(* IEC 61131-3 sources: 2026_Projet_YGO_ExcavatriceDragage/CODE_BACKUP/CODE_20260807_v0.5.25/JOYSTICK, 4 files *)

(* ---- ST_Joystick_AxisCmd.st ---- *)
(* ═══════════════════════════════════════════════════════════════
   🕹️ ST_Joystick_AxisCmd — Consigne d'axe normalisée (sortie FB_Joystick)
   ───────────────────────────────────────────────────────────────
   📄 Doc métier : DOC/AF_Partie-08_Fonction_Joystick_v2.0.md
                   DOC/AF_Partie-03_Contrats_Composants_v2.1.md
   🎯 4 champs exactement :
      - Enable    : Autorisation globale du pipeline
      - StartStop : RAMPE (TRUE = accélération, FALSE = décélération normale)
      - SpeedRef  : Consigne vitesse signée (-100.0 .. +100.0 %)
      - Direction : Sens d'axe (-1 = Rev, 0 = Neutre, +1 = Fwd)
   ═══════════════════════════════════════════════════════════════ *)

TYPE ST_Joystick_AxisCmd :
STRUCT
    Enable      : BOOL;   // Autorisation FB (FALSE = neutralisation, sorties coupées)
    StartStop   : BOOL;   // TRUE = rampe accélération, FALSE = rampe décélération normale
    SpeedRef    : REAL;   // Consigne vitesse SIGNÉE -100..+100 % (signe = sens, cohérent avec Direction)
    Direction   : INT;    // -1 = Rev, 0 = Neutre, +1 = Fwd
END_STRUCT
END_TYPE

(* ---- FB_AxisScale.st ---- *)
(* ═══════════════════════════════════════════════════════════════
   📐 FB_AxisScale — Mise à l'échelle d'un axe joystick Hall
   ───────────────────────────────────────────────────────────────
   📄 Extrait depuis le projet CODESYS (Device.export, JOYSTICK/)
   🎯 Normalise une valeur brute (0..10000) par rapport au neutre calibré
      et applique une zone morte en unités brutes (compte ADC, pas en %).
   Sortie : OutPct ∈ [-100.0 .. +100.0] (0.0 si dans la deadband)
   🔧 2026-08-07 (demande client) : Deadband (REAL, %) → DeadbandRaw (INT, compte brut 0..10000).
      Raison : plus simple à régler directement depuis le bruit mesuré au neutre (ex: ±200 sur le
      terrain → DeadbandRaw=300 avec marge), sans recalculer un % à chaque calibration.
   ═══════════════════════════════════════════════════════════════
   📄 Docs : DOC/AF_Partie-08_Fonction_Joystick_v2.0.md
*)

FUNCTION_BLOCK FB_AxisScale
VAR_INPUT
    /// Valeur brute (0..10000)
    RawIn   : INT;
    /// Point milieu calibré
    Neutral : INT;
    /// Zone morte en unités brutes (compte ADC, ex: 300 sur plage 0..10000)
    DeadbandRaw : INT;
END_VAR
VAR_OUTPUT
    /// Valeur finale (-100.0..100.0)
    OutPct : REAL;
END_VAR
VAR
    Delta : REAL;
END_VAR

IF RawIn >= Neutral THEN
    Delta := INT_TO_REAL(10000 - Neutral);
    IF Delta > 0.0 THEN
        OutPct := (INT_TO_REAL(RawIn - Neutral) / Delta) * 100.0;
    ELSE
        OutPct := 0.0;
    END_IF;
ELSE
    Delta := INT_TO_REAL(Neutral);
    IF Delta > 0.0 THEN
        OutPct := (INT_TO_REAL(RawIn - Neutral) / Delta) * 100.0;
    ELSE
        OutPct := 0.0;
    END_IF;
END_IF;

IF ABS(RawIn - Neutral) <= DeadbandRaw THEN
    OutPct := 0.0;
END_IF;

// 🛡️ Limitation de plage : une valeur brute hors plage nominale ne doit jamais
// produire une consigne supérieure à ±100 %. Ce garde-fou protège les
// consommateurs en aval, notamment la translation M3.
OutPct := LIMIT(-100.0, OutPct, 100.0);

(* ---- FB_Filter_PT1.st ---- *)
(* ═══════════════════════════════════════════════════════════════
   🔁 FB_Filter_PT1 — Filtre passe-bas premier ordre (PT1 numérique)
   ───────────────────────────────────────────────────────────────
   📄 Extrait depuis le projet CODESYS (Device.export, JOYSTICK/)
   🎯 Filtre exponentiel discret : y[k] = α·x[k] + (1-α)·y[k-1]
      où α = CycleTimeS / (T + CycleTimeS), T = TimeConst en secondes.
   ⚠️ Si TimeConst = 0 ou CycleTimeS = 0, sortie = entrée (pass-through).
   ═══════════════════════════════════════════════════════════════
   📄 Docs : DOC/AF_Partie-08_Fonction_Joystick_v2.0.md
*)

FUNCTION_BLOCK FB_Filter_PT1
VAR_INPUT
    /// Consigne brute entrée
    ValueIn    : REAL;
    /// Constante de temps du filtre
    TimeConst  : TIME;
    /// Temps de cycle réel en secondes
    CycleTimeS : REAL;
END_VAR
VAR_OUTPUT
    /// Consigne filtrée sortie
    ValueOut : REAL;
END_VAR
VAR
    T     : REAL;
    Alpha : REAL;
END_VAR

T := TIME_TO_REAL(TimeConst) / 1000.0; // ms → s

IF T <= 0.0 OR CycleTimeS <= 0.0 THEN
    ValueOut := ValueIn;
ELSE
    Alpha    := CycleTimeS / (T + CycleTimeS);
    ValueOut := Alpha * ValueIn + (1.0 - Alpha) * ValueOut;
END_IF;

(* ---- FB_Joystick.st ---- *)
(* ═══════════════════════════════════════════════════════════════
   🕹️ FB_Joystick — Acquisition & traitement Hall (Homme-mort ISO 13850)
   ───────────────────────────────────────────────────────────────
   📄 Doc métier : DOC/AF_Partie-08_Fonction_Joystick_v2.0.md
                   DOC/AF_Partie-03_Contrats_Composants_v2.1.md
   🎯 Rôle : Acquisition 2 axes Hall + bouton homme-mort normatif.
      Pipeline par axe : FB_AxisScale → FB_Filter_PT1 → Homme-Mort → ST_Joystick_AxisCmd.
      Les rampes d'accélération/décélération sont gérées exclusivement par les
      FB de mouvement aval (FB_Winch, FB_Translation), hors de ce bloc.
    🔒 Bouton homme-mort :
       - Armement au neutre strict (ScaleX/Y.OutPct = 0.0).
       - Consentement au démarrage : mouvement libre SANS surveillance du bouton
         (défaut, DeadmanReconfEnable := FALSE). Optionnel : reconfirmation périodique
         en mouvement (délai DeadmanRearmTimeout) si DeadmanReconfEnable := TRUE.
       - Désarmement sur maintien au neutre (durée NeutralHoldTime) + gate/mode/fin benne.
   📤 Produit AxisCmdX, AxisCmdY, et signaux de diagnostic/miroir.
   ═══════════════════════════════════════════════════════════════ *)

// === DECLARATION (à coller dans la partie déclaration du POU FB_Joystick) ===

FUNCTION_BLOCK FB_Joystick
VAR_INPUT
    Enable          : BOOL;       // Active la logique
    Reset           : BOOL;       // Acquittement défaut
    PowerContactorEngaged : BOOL;       // Conditions globales OK (chaîne AU réarmée)
    Mode            : E_Mode;     // Changement de mode désarme le homme-mort
    BenneBusy       : BOOL;       // Fin de cycle benne (front descendant) désarme le homme-mort
    PreserveArmingAfterBucket : BOOL; // TRUE uniquement pendant fermeture ExtractionSequence : enchaînement palier 1 autorisé
    BusCanOpenOP    : ST_Diag_Device;       // État présence nœud CAN
    JoystickOP      : ST_Diag_Device;       // Mode esclave CANopen actif
    RawX            : INT;        // Valeur brute axe X
    RawY            : INT;        // Valeur brute axe Y
    RawButton       : BOOL;       // État brut bouton
    BtnCalibrate    : BOOL;       // Demande de recalage neutre
    InvertX         : BOOL := FALSE;
    InvertY         : BOOL := FALSE;
    DeadbandRaw     : INT := 300;    // 🔧 2026-08-07 (demande client) : zone morte en compte brut ADC (0..10000), remplace l'ancien % — mesure terrain bruit neutre ±200, marge à ±300
    FilterTime      : TIME := TIME#0ms;
    DeadmanRearmTimeout : TIME := T#10S; // Délai max entre 2 appuis en mouvement (si reconfirmation activée)
    NeutralHoldTime     : TIME := T#100MS; // Temps continu au neutre avant désarmement (100 ms)
    DeadmanArmHoldTime  : TIME := T#100MS; // 🆕 2026-08-07 : Temps d'appui continu avant armement (indépendant position axes)
    DeadmanArmGraceTime : TIME := T#3S;    // 🆕 2026-08-07 : Délai après armement avant que le désarmement "neutre tenu" (NeutralHoldTime) puisse s'appliquer — laisse le temps de sortir de la zone morte après un appui au centre
    DeadmanReconfEnable : BOOL := FALSE; // 🆕 2026-08-03 : FALSE = bouton = consentement au démarrage (mouvement libre, défaut cible) ; TRUE = reconfirmation périodique en mouvement (comportement historique)
END_VAR
VAR_OUTPUT
    Ready           : BOOL;       // Prêt à commuter
    Busy            : BOOL;       // Traitement en cours
    Done            : BOOL;       // Données valides dispo
    Error           : BOOL;       // Présence anomalie
    ErrorId         : WORD;       // bit0: "Échec calibration Joystick" - Valeurs RawX/Y hors plage lors du recalage
    AxisCmdX        : ST_Joystick_AxisCmd; // Sortie normalisée X
    AxisCmdY        : ST_Joystick_AxisCmd; // Sortie normalisée Y
    Button          : BOOL;       // Bouton filtré
    NeutralXAct     : INT;        // Point neutre X actuel pour IHM/Test
    NeutralYAct     : INT;        // Point neutre Y actuel pour IHM/Test
    // 🆕 Miroirs directs (maintenance) — mêmes valeurs que AxisCmdX/Y.SpeedRef/.Direction,
    // exposés à plat pour lecture immédiate en vue instance CODESYS (pas de dépliage struct).
    SpeedXPct       : REAL;       // Consigne vitesse axe X en % SIGNÉE (-100..+100), miroir AxisCmdX.SpeedRef
    DirectionX      : INT;        // Sens axe X (-1=Rev/0=Neutre/+1=Fwd), miroir AxisCmdX.Direction
    SpeedYPct       : REAL;       // Consigne vitesse axe Y en % SIGNÉE (-100..+100), miroir AxisCmdY.SpeedRef
    DirectionY      : INT;        // Sens axe Y (-1=Rev/0=Neutre/+1=Fwd), miroir AxisCmdY.Direction
    DeadmanArmed    : BOOL;       // 🆕 Geste armé (bouton appuyé au neutre) — IHM/diagnostic
    AtNeutral       : BOOL;       // 🆕 2026-08-07 : TRUE si les 2 axes sont en zone morte (position centrale) — IHM/diagnostic
END_VAR
VAR_IN_OUT
    NeutralXMem     : INT; // Point neutre X persistant global
    NeutralYMem     : INT; // Point neutre Y persistant global
END_VAR
VAR
    CycleTimeCalc   : FB_CycleTime;
    ScaleX          : FB_AxisScale;
    ScaleY          : FB_AxisScale;
    FilterX         : FB_Filter_PT1;
    FilterY         : FB_Filter_PT1;
    CmdXVal         : REAL;
    CmdYVal         : REAL;
    LastCalibrate   : BOOL;
    ResetEdge       : R_TRIG;
    DeadmanEdge     : R_TRIG;
    DeadmanTimer    : TON;
    NeutralHoldTimer: TON;
    DeadmanArmTimer : TON;
    DeadmanArmPending : BOOL;
    DeadmanArmGraceTimer : TON;
    LastMode        : E_Mode;
    BenneBusyFallEdge : F_TRIG;
END_VAR

// === IMPLEMENTATION (à coller dans le corps ST du POU FB_Joystick) ===

// 🛑 1. GATE (Sécurités et coupures prioritaires)
IF NOT Enable OR NOT PowerContactorEngaged OR NOT BusCanOpenOP.Operational OR NOT JoystickOP.Operational THEN
    Ready := FALSE; Busy := FALSE; Done := FALSE;
    AxisCmdX.Enable := FALSE; AxisCmdX.StartStop := FALSE; AxisCmdX.SpeedRef := 0.0; AxisCmdX.Direction := 0;
    AxisCmdY.Enable := FALSE; AxisCmdY.StartStop := FALSE; AxisCmdY.SpeedRef := 0.0; AxisCmdY.Direction := 0;
    SpeedXPct := 0.0; DirectionX := 0;
    SpeedYPct := 0.0; DirectionY := 0;
    Button := FALSE;
    AtNeutral := TRUE;   // 🆕 2026-08-07 — pas de commande possible pendant la neutralisation
    DeadmanArmed := FALSE;   // 🆕 Désarmé sur toute neutralisation — nouvel appui au neutre exigé
    DeadmanArmPending := FALSE;   // 🆕 2026-08-07 — annule toute tentative d'armement en cours
    DeadmanTimer(IN := FALSE, PT := DeadmanRearmTimeout);   // 🆕 2026-07-03decies — pas d'accumulation à froid
    NeutralHoldTimer(IN := FALSE, PT := NeutralHoldTime);   // 🆕 2026-07-03duodecies — idem
    DeadmanArmTimer(IN := FALSE, PT := DeadmanArmHoldTime);   // 🆕 2026-08-07 — idem
    DeadmanArmGraceTimer(IN := FALSE, PT := DeadmanArmGraceTime);   // 🆕 2026-08-07 — idem
    NeutralXAct := NeutralXMem;
    NeutralYAct := NeutralYMem;
    LastMode := Mode;   // 🆕 REX 2026-07-08 — pas de faux changement détecté à la réactivation
    RETURN;
END_IF;

Ready := TRUE; Busy := TRUE;

// 🔑 2. RESET DÉFAUT (front + cause disparue, Partie3 §5)
ResetEdge(CLK := Reset);
IF ResetEdge.Q AND (RawX >= 2000 AND RawX <= 8000 AND RawY >= 2000 AND RawY <= 8000) THEN
    ErrorId := ErrorId AND 16#FFFE;
END_IF;

// 📥 3. ACQUISITION TIMING & BOUTON
CycleTimeCalc();
Button := RawButton;

// 🎯 4. CALIBRATION DYNAMIQUE (Zone RETAIN)
IF BtnCalibrate AND NOT LastCalibrate THEN
    IF RawX >= 2000 AND RawX <= 8000 AND RawY >= 2000 AND RawY <= 8000 THEN
        NeutralXMem := RawX;
        NeutralYMem := RawY;
    ELSE
        // Un seul bit pour une seule cause (Partie3 §3)
        ErrorId := ErrorId OR 16#0001;
    END_IF;
END_IF;
Error := (ErrorId <> 16#0000);
LastCalibrate := BtnCalibrate;

// 🧮 4bis. MISE À L'ÉCHELLE (avant homme-mort — le neutre s'évalue sur les 2 axes déjà deadbandés)
ScaleX(RawIn := RawX, Neutral := NeutralXMem, DeadbandRaw := DeadbandRaw);
ScaleY(RawIn := RawY, Neutral := NeutralYMem, DeadbandRaw := DeadbandRaw);
AtNeutral := (ScaleX.OutPct = 0.0) AND (ScaleY.OutPct = 0.0);   // 🆕 2026-08-07 : IHM/diagnostic — position centrale (zone morte)

// 4ter-bis. CHANGEMENT DE MODE : désarme le homme-mort dès que Mode change
// (MAINT_N1/N2/SEMI_AUTO/AUTO). Évite qu'une commande en cours traverse le changement
// de mode et soit réinterprétée soudainement. Repassage par le neutre + nouvel appui exigé.
IF Mode <> LastMode THEN
    DeadmanArmed := FALSE;
    DeadmanArmPending := FALSE;   // 🆕 2026-08-07 — nouvel appui exigé après changement de mode
END_IF;
LastMode := Mode;

// 4ter-ter. FIN DE CYCLE BENNE : désarmement général pour qu'une fermeture manuelle
// ne démarre jamais M1/M2 par surprise. Exception : ExtractionSequence garde l'armement
// pendant sa fermeture (enchaînement palier 1 sous ses propres interlocks synchro/position).
BenneBusyFallEdge(CLK := BenneBusy);
IF BenneBusyFallEdge.Q AND NOT PreserveArmingAfterBucket THEN
    DeadmanArmed := FALSE;
    DeadmanArmPending := FALSE;   // 🆕 2026-08-07 — nouvel appui exigé après fin de cycle benne
END_IF;

// 4ter. BOUTON HOMME-MORT — armement par MAINTIEN (DeadmanArmHoldTime), indépendant de la
// position des axes pendant l'appui.
// 🔧 2026-08-07 (retour terrain) : l'ancien armement ("front bouton" ET "axes strictement à
// 0.0 sur le MÊME scan") échouait dès que l'opérateur poussait le joystick quelques ms après
// avoir appuyé — trop contraignant en pratique (le geste naturel "j'appuie PUIS je pousse" ratait
// systématiquement la fenêtre d'un seul scan). Nouvelle séquence : appui (front) → maintien
// DeadmanArmHoldTime (100 ms) → armé, quelle que soit la position des axes durant ce maintien.
// Relâchement AVANT la fin du maintien = tentative annulée (DeadmanArmPending retombe), un
// nouvel appui (front) est requis — pas d'armement différé "surprise" sur un appui prolongé après
// un désarmement (mode/benne/neutre). Sûr même si le joystick est déjà hors zone morte à la fin
// du maintien : les rampes d'accel/décel restent gérées par les FB aval (FB_Winch/FB_Translation,
// cf. §"Rôle" en tête de fichier), donc pas de démarrage brutal possible côté ce FB.
DeadmanEdge(CLK := RawButton);
IF DeadmanEdge.Q THEN
    DeadmanArmPending := TRUE;
END_IF;
IF NOT RawButton THEN
    DeadmanArmPending := FALSE;
END_IF;
DeadmanArmTimer(IN := DeadmanArmPending AND NOT DeadmanArmed, PT := DeadmanArmHoldTime);
IF DeadmanArmTimer.Q THEN
    DeadmanArmed := TRUE;
    DeadmanArmPending := FALSE;
END_IF;

// 🔧 2026-08-06 (retour terrain) : décision 2026-08-03 ("l'opérateur a le temps qu'il veut
// pour démarrer après armement") ANNULÉE explicitement — un armement resté au neutre sans
// mouvement démarré ne désarmait JAMAIS (LeftNeutralSinceArm restait FALSE indéfiniment),
// laissant DeadmanArmed collé à TRUE d'une session à l'autre. Neutre tenu NeutralHoldTime
// désarme désormais TOUJOURS, qu'un mouvement ait été démarré ou non depuis l'armement.
// 🔧 2026-08-07 (retour terrain) : SANS garde-fou, ce désarmement se déclenchait ~100-200ms après
// CHAQUE armement (l'appui se fait typiquement AU neutre depuis le nouvel armement par maintien —
// voir §4ter — donc AtNeutral est déjà vrai dès l'instant où DeadmanArmed passe à TRUE, et
// NeutralHoldTime=100ms est trop court pour laisser le temps de sortir de la zone morte). Ajout
// DeadmanArmGraceTimer (3s) : le désarmement neutre ne peut s'appliquer qu'APRÈS ce délai suivant
// l'armement — le risque du 2026-08-06 (armement collé indéfiniment) reste couvert, juste avec
// une marge de départ au lieu de 100ms. Aucun risque moteur pendant la grâce : au neutre,
// CmdXVal/CmdYVal restent à 0 (deadband), armé ou non.
DeadmanArmGraceTimer(IN := DeadmanArmed, PT := DeadmanArmGraceTime);
NeutralHoldTimer(IN := DeadmanArmed AND AtNeutral AND DeadmanArmGraceTimer.Q,
                 PT := NeutralHoldTime);
IF NeutralHoldTimer.Q THEN
    DeadmanArmed := FALSE;      // Neutre tenu assez longtemps (après la grâce) = désarmement
END_IF;

// 4quater. RECONFIRMATION PÉRIODIQUE (optionnelle) — activée uniquement si DeadmanReconfEnable := TRUE.
// 🆕 2026-08-03 : par défaut FALSE → bouton = CONSENTEMENT AU DÉMARRAGE : une fois armé, le mouvement
// est libre SANS surveillance du bouton ; seuls gate/mode/fin benne/neutre 500ms désarment.
// ⚠️ CORRECTIF (garde-fou si réactivé) : le 1er jet ne détectait qu'un FRONT (`DeadmanEdge.Q`) — un
// opérateur qui MAINTIENT le bouton enfoncé en continu (réflexe naturel homme-mort) ne générait
// plus jamais de front après le 1er appui → désarmement surprise au bout de 3s MALGRÉ la présence
// continue. Corrigé : `NOT RawButton` (niveau, pas front) — maintenir OU réappuyer dans le délai
// remettent tous les deux `IN` à FALSE (TON.ET repart de 0), seul un RELÂCHEMENT PROLONGÉ désarme.
DeadmanTimer(IN := DeadmanReconfEnable AND DeadmanArmed
                   AND NOT AtNeutral AND NOT RawButton,
             PT := DeadmanRearmTimeout);
IF DeadmanTimer.Q THEN
    DeadmanArmed := FALSE;      // Pas de reconfirmation dans le délai → désarmement (décélération sûre)
END_IF;

// 🕹️ 5. PIPELINE TRAITEMENT — AXE X
IF InvertX THEN
    FilterX(ValueIn := -ScaleX.OutPct, TimeConst := FilterTime, CycleTimeS := CycleTimeCalc.CycleTimeS);
ELSE
    FilterX(ValueIn := ScaleX.OutPct, TimeConst := FilterTime, CycleTimeS := CycleTimeCalc.CycleTimeS);
END_IF;

// Consigne forcée à 0.0 tant que le geste n'est pas armé (homme-mort)
CmdXVal := SEL(DeadmanArmed, 0.0, FilterX.ValueOut);

// Mapping Sortie Standardisée Axe X
AxisCmdX.Enable := TRUE;
AxisCmdX.SpeedRef := CmdXVal;
AxisCmdX.StartStop := (ABS(CmdXVal) > 0.1);

IF CmdXVal > 0.1 THEN
    AxisCmdX.Direction := 1;
ELSIF CmdXVal < -0.1 THEN
    AxisCmdX.Direction := -1;
ELSE
    AxisCmdX.Direction := 0;
    AxisCmdX.SpeedRef := 0.0;
END_IF;

// Miroirs maintenance
SpeedXPct := AxisCmdX.SpeedRef;
DirectionX := AxisCmdX.Direction;

// 🕹️ 6. PIPELINE TRAITEMENT — AXE Y
IF InvertY THEN
    FilterY(ValueIn := -ScaleY.OutPct, TimeConst := FilterTime, CycleTimeS := CycleTimeCalc.CycleTimeS);
ELSE
    FilterY(ValueIn := ScaleY.OutPct, TimeConst := FilterTime, CycleTimeS := CycleTimeCalc.CycleTimeS);
END_IF;

// Consigne forcée à 0.0 tant que le geste n'est pas armé (homme-mort)
CmdYVal := SEL(DeadmanArmed, 0.0, FilterY.ValueOut);

// Mapping Sortie Standardisée Axe Y
AxisCmdY.Enable := TRUE;
AxisCmdY.SpeedRef := CmdYVal;
AxisCmdY.StartStop := (ABS(CmdYVal) > 0.1);

IF CmdYVal > 0.1 THEN
    AxisCmdY.Direction := 1;
ELSIF CmdYVal < -0.1 THEN
    AxisCmdY.Direction := -1;
ELSE
    AxisCmdY.Direction := 0;
    AxisCmdY.SpeedRef := 0.0;
END_IF;

// Miroirs maintenance
SpeedYPct := AxisCmdY.SpeedRef;
DirectionY := AxisCmdY.Direction;

// 📤 7. VALIDATION DES SORTIES ÉTAT
NeutralXAct := NeutralXMem;
NeutralYAct := NeutralYMem;
Done := NOT Error;
